SUBAPPLICATION Uebung_162b_AX (* Übung zu DS18B20: zwei Sensoren, einer per ROM-Code festgehalten *)
  (* Standard: 61499-2; Description: Copyright (c) 2026 Meisterschulen am Ostbahnhof This program and the accompanying materials are made available under the terms of the Eclipse Public License 2.0 which is available at https://www.eclipse.org/legal/epl-2.0/ SPDX-License-Identifier: EPL-2.0 *)
  (* Version 1.0, 2026-11-26, Franz Höpfinger, Meisterschulen am Ostbahnhof, initial API and implementation and/or initial documentation *)
  PACKAGE Uebungen;
  IMPORT logiBUS::io::DQ::logiBUS_DO::Output_Q1;
  IMPORT logiBUS::io::DQ::logiBUS_DO::Output_Q2;
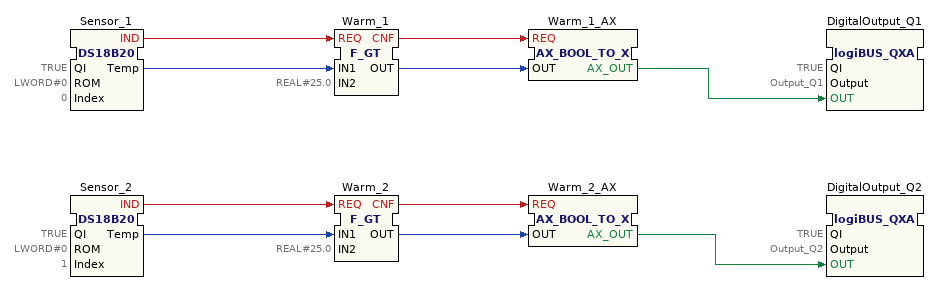
  (* Zwei Temperatursensoren DS18B20 am selben 1-Wire-Bus (Trainer20: GPIO3, bis zu 8 Sensoren). Sensor_1 nimmt den ersten Sensor der Suche (Index 0), Sensor_2 den zweiten (Index 1). Q1/Q2 an = wärmer als 25 °C. Die Suchreihenfolge hängt am ROM-Code. Kommt ein Sensor dazu, kann sich die Zuordnung ändern. Festhalten: Sensor_2.ROMO im Watch ablesen und als ROM (LWORD#16#...) bei Sensor_2 eintragen. Dann zählt Index nicht mehr. Watch: Temp, QO, STATUS, ROMO je Sensor. *)
  FBS
    Sensor_1 : logiBUS::onewire::DS18B20(QI := TRUE, ROM := LWORD#0, Index := 0); (* erster Sensor in Suchreihenfolge *)
    Warm_1 : iec61131::comparison::F_GT(IN2 := REAL#25.0); (* Sensor 1 über 25 °C? *)
    Warm_1_AX : adapter::conversion::unidirectional::AX_BOOL_TO_X;
    DigitalOutput_Q1 : logiBUS::io::DQ::logiBUS_QXA(QI := TRUE, Output := Output_Q1); (* an = Sensor 1 wärmer als 25 °C *)
    Sensor_2 : logiBUS::onewire::DS18B20(QI := TRUE, ROM := LWORD#0, Index := 1); (* Index 1, oder ROMO als ROM eintragen *)
    Warm_2 : iec61131::comparison::F_GT(IN2 := REAL#25.0); (* Sensor 2 über 25 °C? *)
    Warm_2_AX : adapter::conversion::unidirectional::AX_BOOL_TO_X;
    DigitalOutput_Q2 : logiBUS::io::DQ::logiBUS_QXA(QI := TRUE, Output := Output_Q2); (* an = Sensor 2 wärmer als 25 °C *)
  END_FBS
  EVENT_CONNECTIONS
    Sensor_1.IND TO Warm_1.REQ;
    Warm_1.CNF TO Warm_1_AX.REQ;
    Sensor_2.IND TO Warm_2.REQ;
    Warm_2.CNF TO Warm_2_AX.REQ;
  END_CONNECTIONS
  DATA_CONNECTIONS
    Sensor_1.Temp TO Warm_1.IN1;
    Warm_1.OUT TO Warm_1_AX.OUT;
    Sensor_2.Temp TO Warm_2.IN1;
    Warm_2.OUT TO Warm_2_AX.OUT;
  END_CONNECTIONS
  ADAPTER_CONNECTIONS
    Warm_1_AX.AX_OUT TO DigitalOutput_Q1.OUT;
    Warm_2_AX.AX_OUT TO DigitalOutput_Q2.OUT;
  END_CONNECTIONS
END_SUBAPPLICATION
